Fanuc KAREL source: KB00013.KL

PROGRAM KB00013
%NOLOCKGROUP
%ENVIRONMENT FLBT
VAR
  P1: FILE
  P2: INTEGER
  P3: INTEGER
BEGIN
  P2 = 1
  P3 = 1
  BYTES_AHEAD(P1, P2, P3)
END KB00013
